Staubli VAL3: Project.pjx

--- Project.pjx ---
parameters version=s6.8 stackSize=5000 millimeterUnit=true
program file=start.pgx
program file=stop.pgx
program file=feedCylinder.pgx
program file=pickPlaceCylinder.pgx
program file=pickInsertPiston.pgx
program file=placeInMatrix.pgx
data file=Data.dtx
data file=io.dtx

--- Data.dtx ---


--- start.pgx ---
program start()
// Lab2B - Level 3: Continuous assembly with piston presence sensing and matrix palletizing.
begin
  userPage()
  cls()
  putln("====================================")
  putln("  Lab2B - LEVEL 3 (TX60 Assembly)   ")
  putln("====================================")

  // Initialize state and dispenser actuator
  nPistonIdx = 0
  bOut10 = false
  open(tLateral)

  for nCycle = 0 to (nTotalCycles - 1)
    putln("")
    putln("--- CYCLE " + toString("1.0", nCycle + 1) + " / " + toString("1.0", nTotalCycles) + " ---")

    // 1. Ensure red cylinder is fed in dispenser
    call feedCylinder()

    // 2. Pick cylinder and place in assembling station
    call pickPlaceCylinder()

    // 3. Scan piston source with sensor bIn0, pick piston and insert
    call pickInsertPiston()

    // 4. Pick assembled unit and place in Assembled Matrix
    call placeInMatrix(nCycle)
  endFor

  putln("")
  putln("Returning to safe home posture...")
  movej(jStart, flange, mNomSpeed)
  waitEndMove()
  putln("LEVEL 3 COMPLETED SUCCESSFULLY!")
end

--- feedCylinder.pgx ---
program feedCylinder()
// Controls the cylinder dispenser pneumatic actuator and verifies part presence.
begin
  putln("[1/4] Checking cylinder dispenser...")

  while bIn2 == false
    putln("  -> No cylinder ready. Actuating feeder...")

    // Guarantee actuator starts fully contracted
    if bIn15 == false
      bOut10 = false
      wait(bIn15 == true)
    endIf

    // Extend pneumatic piston to push cylinder out
    bOut10 = true
    wait(bIn14 == true)
    delay(0.2)

    // Contract pneumatic piston back to rest
    bOut10 = false
    wait(bIn15 == true)
    delay(0.2)

    // If still empty, magazine tube needs refilling
    if bIn2 == false
      putln("  [!] Magazine empty! Refill red cylinders...")
      delay(2.0)
    endIf
  endWhile

  putln("  -> Red cylinder ready at pick position.")
end

--- pickInsertPiston.pgx ---
program pickInsertPiston()
// Scans 2x4 Piston Source using tool sensor bIn0, picks available piston, and inserts it.
  local num nRow
  local num nCol
  local point pCurPick
  local point pCurCheck
  local point pCurApp
begin
  putln("[3/4] Scanning piston source (bIn0)...")
  open(tTip)
  bPistonFound = false

  while !bPistonFound
    // Wrap around if all 8 slots were scanned without finding a piston
    if nPistonIdx >= (nPistonRows * nPistonCols)
      putln("  [!] Tray empty! Refill pistons in source...")
      nPistonIdx = 0
      delay(2.0)
    endIf

    // Compute (row, col) in 2x4 Piston Source grid
    nRow = roundDown(nPistonIdx / nPistonCols)
    nCol = nPistonIdx - (nRow * nPistonCols)

    pCurPick = pPistonBase
    pCurPick.trsf.x = pPistonBase.trsf.x + (nCol * nPistonStepX)
    pCurPick.trsf.y = pPistonBase.trsf.y + (nRow * nPistonStepY)

    pCurCheck = appro(pCurPick, trPistonSensor)
    pCurApp = appro(pCurPick, trPistonAppro)

    // Move above slot and check presence sensor bIn0
    movej(pCurApp, tTip, mNomSpeed)
    waitEndMove()
    movel(pCurCheck, tTip, mNomSpeed)
    waitEndMove()
    delay(0.15)

    if bIn0 == true
      bPistonFound = true
      putln("  -> Piston FOUND at [" + toString("1.0", nRow) + "," + toString("1.0", nCol) + "]")

      movel(pCurPick, tTip, mInsertSpeed)
      waitEndMove()
      close(tTip)

      movel(pCurApp, tTip, mNomSpeed)
      waitEndMove()
    else
      putln("  -> Slot [" + toString("1.0", nRow) + "," + toString("1.0", nCol) + "] EMPTY, skipping...")
      movel(pCurApp, tTip, mNomSpeed)
      waitEndMove()
    endIf

    // Advance index for next check/cycle
    nPistonIdx = nPistonIdx + 1
  endWhile

  // Insert piston into cylinder at assembling station
  putln("  -> Inserting piston into cylinder...")
  movej(pInsertApproach, tTip, mNomSpeed)
  waitEndMove()
  movel(pInsert, tTip, mInsertSpeed)
  waitEndMove()
  open(tTip)

  movel(pInsertApproach, tTip, mNomSpeed)
  waitEndMove()
end

--- pickPlaceCylinder.pgx ---
program pickPlaceCylinder()
// Picks red cylinder from dispenser and places it in the assembling station.
begin
  putln("[2/4] Transferring red cylinder to station...")
  open(tLateral)

  // Safe joint transit to avoid wrist/elbow flip
  movej(jTransCylinder, tLateral, mNomSpeed)
  waitEndMove()

  // Pick from dispenser
  movej(pCylApproach, tLateral, mNomSpeed)
  waitEndMove()
  movel(pCylPick, tLateral, mInsertSpeed)
  waitEndMove()
  close(tLateral)

  movel(pCylApproach, tLateral, mNomSpeed)
  waitEndMove()

  // Place in assembling station
  movej(pAsmApproach, tLateral, mNomSpeed)
  waitEndMove()
  movel(pAsmCylinder, tLateral, mInsertSpeed)
  waitEndMove()
  open(tLateral)

  movel(pAsmApproach, tLateral, mNomSpeed)
  waitEndMove()
end

--- placeInMatrix.pgx ---
program placeInMatrix(num nSlotIdx (byVal=true))
// Picks assembled unit from station and places it into the corresponding fMatrix slot.
  local num nRow
  local num nCol
  local point pCurPlace
  local point pCurApp
begin
  putln("[4/4] Placing assembly into matrix...")
  open(tLateral)

  // Pick assembled unit from assembling station
  movej(pAsmApproach, tLateral, mNomSpeed)
  waitEndMove()
  movel(pAsmCylinder, tLateral, mInsertSpeed)
  waitEndMove()
  close(tLateral)

  movel(pAsmApproach, tLateral, mNomSpeed)
  waitEndMove()

  // Compute (row, col) in 2x4 Assembled Matrix
  nRow = roundDown(nSlotIdx / nMatrixCols)
  nCol = nSlotIdx - (nRow * nMatrixCols)

  pCurPlace = pMatrixBase
  pCurPlace.trsf.x = pMatrixBase.trsf.x + (nCol * nMatrixStepX)
  pCurPlace.trsf.y = pMatrixBase.trsf.y + (nRow * nMatrixStepY)
  pCurApp = appro(pCurPlace, trMatrixAppro)

  putln("  -> Target matrix slot [" + toString("1.0", nRow) + "," + toString("1.0", nCol) + "]")

  movej(pCurApp, tLateral, mNomSpeed)
  waitEndMove()
  movel(pCurPlace, tLateral, mInsertSpeed)
  waitEndMove()
  open(tLateral)

  movel(pCurApp, tLateral, mNomSpeed)
  waitEndMove()
end

--- stop.pgx ---
program stop()
// Safe stop routine: halts motion and resets feeder valve without dropping held parts.
begin
  resetMotion()
  bOut10 = false
  putln("Lab2B stopped safely - gripper state preserved")
end
